{attribute 'qualified_only'}
{attribute 'strict'}
TYPE E_OwnerDevice :
(
	NotDefined := 0,
	Tank1,
	Tank2,
	Tank3,
	Tank4,
	common //last
);
END_TYPE

(* stored: Version 1.1.0.1, ProductVersion 3.1.4024.12
   DUT E_OwnerDevice: Id {22e48fdb-8d6e-4e9b-bfa5-d24f2ffac593} *)
